// Function block for calculating the sum of two values
FUNCTION_BLOCK FB_Sum
VAR_INPUT
	var1: UINT;    // variable 1
	var2: UINT;    // variable 2
END_VAR
VAR_OUTPUT
	result : UINT; // result
END_VAR

// Calculation of the sum of two values; an error has been deliberately included in this example
result := var1 - var2;

END_FUNCTION_BLOCK

(* stored: Version 1.1.0.1, ProductVersion 3.1.4026.18
   POU FB_Sum: Id {7e3cb313-c37d-401b-91eb-437d061cc677}, SpecialFunc None *)
